Fanuc KAREL source: KT00505.KL

PROGRAM KT00505
%NOLOCKGROUP
VAR
  P1: XYZWPR
  P2: XYZWPREXT
  OUT: XYZWPR
BEGIN
  P1.X = 1.0
    P2.Y = 2.0
  OUT = P1 : P2
END KT00505
